Fanuc KAREL source: ka00055.KL

PROGRAM KA00055
%STACKSIZE=65535
%PRIORITY=65535
%NOLOCKGROUP
VAR
SRC : POSITION
DST : XYZWPREXT
BEGIN
-- UNSAFE_SOURCE_IR line 7: DST = convert_position_to_xyzwprext(SRC)
END KA00055
